// ---- POUs/POUs/FB/FB_Station05_Tear.TcPOU
FUNCTION_BLOCK FB_Station05_Tear EXTENDS FB_RollerConveyor
// =============================================================
// STACJA 5 - TEST WYTRZYMALOSCI NA ROZRYWANIE
// =============================================================
//
// Transporter rolkowy plus mechanika testu: blokada punktu
// zatrzymania, podnoszone szczeki chwytajace dolne deski
// i szesc silownikow rozrywajacych napierajacych na deski gorne.
//
// -------------------------------------------------------------
// DLACZEGO NIE MA PRZEJAZDU BEZ ZATRZYMANIA
// -------------------------------------------------------------
// Blokada stoi dokladnie w punkcie zatrzymania. Zeby przepuscic
// palete bez postoju, trzeba by ja opuscic ZANIM paleta dojedzie,
// czyli podjac decyzje na podstawie stanu, ktory dopiero ma
// nastapic. Blad w tej decyzji to paleta wjezdzajaca w podniesiona
// blokade z pelna predkoscia.
//
// Dlatego stacja 5 zatrzymuje KAZDA palete, takze odrzucona
// i takze przy wylaczonym tescie - wtedy sekwencja sprowadza sie
// do opuszczenia blokady. W GVL_PERSIST.aConv[5].Cfg nalezy
// ustawic xAllowPassThrough := FALSE.
//
// -------------------------------------------------------------
// KIEDY PODNOSI SIE BLOKADA
// -------------------------------------------------------------
// W chwili, gdy z poprzedniej stacji RUSZA paleta - czyli
// w M_BeginInfeed. Wtedy droga jest wolna na pewno, a czasu na
// ruch jest tyle, ile trwa przejazd miedzy stacjami.
//
// Podnoszenie jej czasowka po zjezdzie poprzedniej palety
// byloby zgadywaniem, czy paleta zeszla juz z blokady.
//
// -------------------------------------------------------------
// PRZEBIEG TESTU
// -------------------------------------------------------------
//   10  czasowka od potwierdzenia palety na blokadzie
//   20  podniesienie szczek
//   30  zamkniecie szczek (3 pary)
//   40  czasowka przed rozrywaniem
//   50  rozrywanie - kazdy silownik badany OSOBNO
//   60  otwarcie szczek
//   70  opuszczenie szczek
//   80  opuszczenie blokady
//   90  koniec
//
// Kazdy silownik rozrywajacy ma wlasny licznik czasu trzymania
// nacisku, bo wszystkie ida z inna predkoscia. Przekroczenie
// progu polozenia = deska odpadla: paleta staje sie NOK i nie
// przechodzi juz zadnych dalszych testow ani etykietowania.
VAR_INPUT

	stIn	: ST_St05_In;

END_VAR
VAR_OUTPUT

	stOut	: ST_St05_Out;

	// Krok sekwencji testu - do podgladu na HMI
	nTestStep		: INT;

	// Ktorego silownika rozrywajacego jeszcze czekamy (0 = zaden)
	nWaitPull		: INT;

	// Wynik dla biezacej palety
	axBoardBroken	: ARRAY[1..6] OF BOOL;

	// Wolna droga dla wjazdu: szczeki otwarte i opuszczone,
	// silowniki rozrywajace wycofane. Blokada NIE jest tu
	// warunkiem - podnosi sie dopiero w chwili wjazdu.
	xEntryReady		: BOOL;

	// Pelne polozenie spoczynkowe, z blokada w gorze
	xHomePosition	: BOOL;

	// Pierwszy silownik zglaszajacy blad i jego przyczyna.
	// nFaultyCyl: 1..3 szczeki, 4 blokada, 5 podnoszenie szczek,
	//             6..11 silowniki rozrywajace 1..6
	nFaultyCyl		: INT;
	eCylAlarm		: E_CylAlarm;

END_VAR
VAR

	pSt				: POINTER TO ST_St05Cfg;

	// Blokada punktu zatrzymania
	fbBlock			: FB_Cylinder;

	// Podnoszenie i opuszczanie szczek
	fbJawLift		: FB_Cylinder;

	// Szczeki - trzy pary, kazda para jeden zawor
	fbJaw			: ARRAY[1..3] OF FB_Cylinder;

	// Silowniki rozrywajace, indeksowane NUMEREM SILOWNIKA
	fbPull			: ARRAY[1..6] OF FB_Cylinder;

	axPullDone		: ARRAY[1..6] OF BOOL;

	tonSeq			: TON;
	tonOpWd			: TON;

	i				: INT;
	xAllJawsOpen	: BOOL;
	xAllJawsClosed	: BOOL;
	xAllPullBack	: BOOL;

END_VAR
VAR CONSTANT

	ST5_IDLE			: INT := 0;
	ST5_DELAY			: INT := 10;
	ST5_JAWLIFT_UP		: INT := 20;
	ST5_JAWS_CLOSE		: INT := 30;
	ST5_SETTLE			: INT := 40;
	ST5_PULL			: INT := 50;
	ST5_JAWS_OPEN		: INT := 60;
	ST5_JAWLIFT_DOWN	: INT := 70;
	ST5_BLOCK_DOWN		: INT := 80;
	ST5_DONE			: INT := 90;

END_VAR

// =============================================================
// CYKL STACJI 5
// =============================================================


// 1. Odswiezenie sprzezen silownikow.
//    Robimy to PRZED sekwencja, zeby decyzja "deska odpadla"
//    zapadala na swiezym odczycie przetwornika.
M_CallCylinders();


// 2. Warstwa transportu - wola M_OperationRequired
//    i M_OperationCycle
SUPER^();


// 3. Sprowadzenie mechaniki do polozenia spoczynkowego,
//    gdy stacja jest pusta
M_HomeCycle();


// 4. Przepisanie cewek na strukture wyjsciowa
M_MapOutputs();

METHOD PUBLIC M_ConfigStation
// Podpiecie nastaw stacji i wszystkich silownikow.
// Wolac raz, przy starcie, PO M_Config klasy bazowej.
VAR_INPUT
	pStCfg		: POINTER TO ST_St05Cfg;

	// Tablica rekordow silownikow - ADR(GVL_PERSIST.aCyl)
	pCylArray	: POINTER TO ARRAY[1..32] OF ST_CylPersist;

	// Pierwszy indeks przydzielony stacji. Stacja zajmuje
	// 11 kolejnych rekordow: szczeki 1..3, blokada,
	// podnoszenie szczek, silowniki rozrywajace 1..6.
	nCylBase	: INT;
END_VAR
VAR
	j			: INT;
END_VAR
pSt := pStCfg;

IF pCylArray = 0 THEN
	RETURN;
END_IF


// Szczeki
FOR j := 1 TO 3 DO
	fbJaw[j].M_Config(
		nId			:= nCylBase + j - 1,
		pPersist	:= ADR(pCylArray^[nCylBase + j - 1])
	);
END_FOR

// Blokada punktu zatrzymania
fbBlock.M_Config(
	nId			:= nCylBase + 3,
	pPersist	:= ADR(pCylArray^[nCylBase + 3])
);

// Podnoszenie szczek
fbJawLift.M_Config(
	nId			:= nCylBase + 4,
	pPersist	:= ADR(pCylArray^[nCylBase + 4])
);

// Silowniki rozrywajace
FOR j := 1 TO 6 DO
	fbPull[j].M_Config(
		nId			:= nCylBase + 4 + j,
		pPersist	:= ADR(pCylArray^[nCylBase + 4 + j])
	);
END_FOR
END_METHOD

METHOD PROTECTED M_CallCylinders
// Wywolanie wszystkich silownikow z ich sygnalami wejsciowymi
// oraz zebranie zbiorczych warunkow mechaniki.
VAR
	j	: INT;
END_VAR
fbBlock(
	eMode		:= eMode,
	xSafetyOK	:= xSafetyOK,
	xSwExtRaw	:= stIn.xBlockUpSw,
	xSwRetRaw	:= stIn.xBlockDownSw
);

fbJawLift(
	eMode		:= eMode,
	xSafetyOK	:= xSafetyOK,
	xSwExtRaw	:= stIn.xJawLiftUpSw,
	xSwRetRaw	:= stIn.xJawLiftDownSw
);


// Para szczek jest otwarta dopiero gdy OBA silowniki
// zglaszaja otwarcie
xAllJawsOpen	:= TRUE;
xAllJawsClosed	:= TRUE;

FOR j := 1 TO 3 DO

	fbJaw[j](
		eMode		:= eMode,
		xSafetyOK	:= xSafetyOK,
		xSwExtRaw	:= FALSE,
		xSwRetRaw	:= stIn.axJawOpenSw[j, 1] AND stIn.axJawOpenSw[j, 2]
	);

	IF NOT fbJaw[j].xRetracted THEN
		xAllJawsOpen := FALSE;
	END_IF

	IF NOT fbJaw[j].xExtended THEN
		xAllJawsClosed := FALSE;
	END_IF

END_FOR


xAllPullBack := TRUE;

FOR j := 1 TO 6 DO

	fbPull[j](
		eMode		:= eMode,
		xSafetyOK	:= xSafetyOK,
		diPosRaw	:= stIn.adiPullPos[j]
	);

	IF NOT fbPull[j].xRetracted THEN
		xAllPullBack := FALSE;
	END_IF

END_FOR


// Wolna droga dla wjazdu. Blokada nie jest tu warunkiem -
// podnosi sie dopiero wtedy, gdy z poprzedniej stacji rusza
// paleta, wiec przy pustej stacji stoi w dole.
xEntryReady := fbJawLift.xRetracted AND xAllJawsOpen AND xAllPullBack;

xHomePosition := xEntryReady AND fbBlock.xExtended;


M_ScanCylinderFaults();
END_METHOD

METHOD PROTECTED M_MapOutputs
VAR
	j	: INT;
END_VAR
stOut.xBlockExtend		:= fbBlock.xCoilExtend;
stOut.xBlockRetract		:= fbBlock.xCoilRetract;

stOut.xJawLiftExtend	:= fbJawLift.xCoilExtend;
stOut.xJawLiftRetract	:= fbJawLift.xCoilRetract;

FOR j := 1 TO 3 DO
	stOut.axJawClose[j] := fbJaw[j].xCoilExtend;
END_FOR

FOR j := 1 TO 6 DO
	stOut.axPullUp[j]	:= fbPull[j].xCoilExtend;
	stOut.axPullDown[j]	:= fbPull[j].xCoilRetract;
END_FOR
END_METHOD

METHOD PROTECTED M_HomeCycle
// Sprowadzenie mechaniki do polozenia gotowosci, gdy stacja
// jest pusta: szczeki otwarte i opuszczone, silowniki
// rozrywajace wycofane.
//
// BLOKADY TU NIE RUSZAMY. Podnosi sie dopiero w chwili, gdy
// z poprzedniej stacji rusza paleta - patrz M_BeginInfeed.
// Podnoszenie jej na czasowke po zjezdzie poprzedniej palety
// oznaczaloby zgadywanie, czy paleta zeszla juz z blokady.
//
// Poza stanem pustym komendy zostaja takie, jakie zostawila
// sekwencja testu.
VAR
	j	: INT;
END_VAR
IF (eState <> NODE_EMPTY) AND (eState <> NODE_INIT) THEN
	RETURN;
END_IF

fbJawLift.M_Retract();

FOR j := 1 TO 3 DO
	fbJaw[j].M_Retract();
END_FOR

FOR j := 1 TO 6 DO
	fbPull[j].M_Retract();
END_FOR
END_METHOD

METHOD PUBLIC M_BeginInfeed
// Poprzednia stacja wlasnie ruszyla z paleta.
//
// To jest moment na podniesienie blokady: droga jest wolna,
// paleta dopiero wjezdza, a czasu na ruch jest tyle, ile trwa
// przejazd miedzy stacjami. Nie zgadujemy niczego czasowka.
VAR_INPUT
	pSource		: POINTER TO FB_TransportNodeBase;
	xNok		: BOOL;
	nLoadId		: UDINT;
END_VAR
SUPER^.M_BeginInfeed(
	pSource	:= pSource,
	xNok	:= xNok,
	nLoadId	:= nLoadId
);

fbBlock.M_Extend();
END_METHOD

METHOD PROTECTED M_ScanCylinderFaults
// Pierwszy silownik w bledzie zostaje wskazany na wyjsciu,
// a stacja idzie w alarm. Kolejne go nie nadpisuja - operator
// ma zobaczyc przyczyne, nie skutek.
VAR
	j	: INT;
END_VAR
IF nFaultyCyl <> 0 THEN
	RETURN;
END_IF

FOR j := 1 TO 3 DO
	IF fbJaw[j].xAlarm AND (nFaultyCyl = 0) THEN
		nFaultyCyl	:= j;
		eCylAlarm	:= fbJaw[j].eAlarm;
	END_IF
END_FOR

IF fbBlock.xAlarm AND (nFaultyCyl = 0) THEN
	nFaultyCyl	:= 4;
	eCylAlarm	:= fbBlock.eAlarm;
END_IF

IF fbJawLift.xAlarm AND (nFaultyCyl = 0) THEN
	nFaultyCyl	:= 5;
	eCylAlarm	:= fbJawLift.eAlarm;
END_IF

FOR j := 1 TO 6 DO
	IF fbPull[j].xAlarm AND (nFaultyCyl = 0) THEN
		nFaultyCyl	:= 5 + j;
		eCylAlarm	:= fbPull[j].eAlarm;
	END_IF
END_FOR

IF nFaultyCyl <> 0 THEN
	M_RaiseAlarm(eNew := ALM_OPERATION_FAILED);
END_IF
END_METHOD

METHOD PUBLIC M_WhyCannotAccept : E_WaitCause
// Warunki klasy bazowej plus wlasne: paleta nie ma prawa
// wjechac, dopoki blokada nie stoi w gorze, a szczeki nie sa
// otwarte i opuszczone.
M_WhyCannotAccept := SUPER^.M_WhyCannotAccept();

IF M_WhyCannotAccept <> WAIT_NONE THEN
	RETURN;
END_IF

IF NOT xEntryReady THEN
	M_WhyCannotAccept := WAIT_STATION_NOT_READY;
END_IF
END_METHOD

METHOD PROTECTED M_OperationRequired : BOOL
// Zawsze TRUE. Nawet paleta odrzucona i nawet przy wylaczonym
// tescie musi sie tu zatrzymac - blokada stoi w punkcie
// zatrzymania i trzeba ja opuscic, zanim paleta pojedzie dalej.
M_OperationRequired := TRUE;
END_METHOD

METHOD PROTECTED M_TestEnabled : BOOL
// Czy dla tej palety w ogole robimy test.
M_TestEnabled := FALSE;

IF pP = 0 THEN
	RETURN;
END_IF

// Operator wylaczyl stacje
IF NOT pP^.Cfg.xStationEnabled THEN
	RETURN;
END_IF

// Paleta juz odrzucona - zadnych dalszych testow
IF pP^.Mem.xLoadNok THEN
	RETURN;
END_IF

M_TestEnabled := TRUE;
END_METHOD

METHOD PROTECTED M_OperationCycle : BOOL
// Sekwencja stacji. Zwraca TRUE, gdy paleta moze jechac dalej.
VAR
	j	: INT;
END_VAR
M_OperationCycle := FALSE;

IF pSt = 0 THEN
	M_RaiseAlarm(eNew := ALM_NOT_CONFIGURED);
	RETURN;
END_IF


// ---------------------------------------------------------
// WATCHDOG CALEJ OPERACJI
// ---------------------------------------------------------

tonOpWd(IN := (nTestStep <> ST5_IDLE), PT := pSt^.tOpWatchdog);

IF tonOpWd.Q THEN
	M_RaiseAlarm(eNew := ALM_OPERATION_FAILED);
	RETURN;
END_IF


CASE nTestStep OF

ST5_IDLE:
	// Start operacji dla nowej palety
	nWaitPull := 0;

	FOR j := 1 TO 6 DO
		axBoardBroken[j]	:= FALSE;
		axPullDone[j]		:= FALSE;
	END_FOR

	tonSeq(IN := FALSE);

	IF M_TestEnabled() THEN
		nTestStep := ST5_DELAY;
	ELSE
		// Bez testu idziemy przez wycofywanie mechaniki, a nie
		// prosto do blokady. Przy pustej stacji te kroki mijaja
		// natychmiast, ale gdy test zostal przerwany w polowie
		// i paleta stala sie NOK - szczeki i silowniki moga byc
		// w dowolnym polozeniu i trzeba je najpierw sciagnac.
		nTestStep := ST5_JAWS_OPEN;
	END_IF


ST5_DELAY:
	tonSeq(IN := TRUE, PT := pSt^.tDetectToLift);

	IF tonSeq.Q THEN
		tonSeq(IN := FALSE);
		nTestStep := ST5_JAWLIFT_UP;
	END_IF


ST5_JAWLIFT_UP:
	fbJawLift.M_Extend();

	IF fbJawLift.xExtended THEN
		nTestStep := ST5_JAWS_CLOSE;
	END_IF


ST5_JAWS_CLOSE:
	FOR j := 1 TO 3 DO
		fbJaw[j].M_Extend();
	END_FOR

	IF xAllJawsClosed THEN
		nTestStep := ST5_SETTLE;
	END_IF


ST5_SETTLE:
	tonSeq(IN := TRUE, PT := pSt^.tJawsToPull);

	IF tonSeq.Q THEN
		tonSeq(IN := FALSE);
		nTestStep := ST5_PULL;
	END_IF


ST5_PULL:
	M_PullCycle();

	IF xAllPullBack AND (nWaitPull = 0) THEN
		nTestStep := ST5_JAWS_OPEN;
	END_IF


ST5_JAWS_OPEN:
	// Silowniki rozrywajace sciagamy takze tutaj - tedy prowadzi
	// droga wyjscia z przerwanego testu
	FOR j := 1 TO 6 DO
		fbPull[j].M_Retract();
	END_FOR

	FOR j := 1 TO 3 DO
		fbJaw[j].M_Retract();
	END_FOR

	IF xAllJawsOpen AND xAllPullBack THEN
		nTestStep := ST5_JAWLIFT_DOWN;
	END_IF


ST5_JAWLIFT_DOWN:
	fbJawLift.M_Retract();

	IF fbJawLift.xRetracted THEN
		nTestStep := ST5_BLOCK_DOWN;
	END_IF


ST5_BLOCK_DOWN:
	fbBlock.M_Retract();

	IF fbBlock.xRetracted THEN
		nTestStep := ST5_DONE;
	END_IF


ST5_DONE:
	// Wyjazd dozwolony dopiero gdy WSZYSTKO jest wycofane
	IF NOT xAllJawsOpen THEN
		RETURN;
	END_IF

	IF NOT fbJawLift.xRetracted THEN
		RETURN;
	END_IF

	IF NOT xAllPullBack THEN
		RETURN;
	END_IF

	IF NOT fbBlock.xRetracted THEN
		RETURN;
	END_IF

	tonOpWd(IN := FALSE);
	nTestStep			:= ST5_IDLE;
	M_OperationCycle	:= TRUE;


ELSE
	nTestStep := ST5_IDLE;

END_CASE
END_METHOD

METHOD PROTECTED M_PullCycle
// Rozrywanie. Kazdy silownik prowadzony OSOBNO - maja rozne
// predkosci, wiec kazdy dochodzi do progu w innej chwili
// i kazdy ma wlasny licznik czasu trzymania nacisku.
VAR
	j	: INT;
END_VAR
nWaitPull := 0;

FOR j := 1 TO 6 DO

	M_PullOne(j := j);

	IF NOT axPullDone[j] THEN
		nWaitPull := j;
	END_IF

END_FOR
END_METHOD

METHOD PROTECTED M_PullOne
// Jeden silownik rozrywajacy.
//
// Kolejnosc warunkow jest istotna: najpierw sprawdzamy, czy
// deska odpadla, i dopiero potem czy nacisk zostal utrzymany.
// Odwrotnie mozna by uznac za dobra deske, ktora wlasnie pekla.
VAR_INPUT
	j	: INT;
END_VAR
// Ten juz zbadany - wraca do bazy
IF axPullDone[j] THEN
	fbPull[j].M_Retract();
	RETURN;
END_IF


// Wysunal sie dalej, niz moglby z cala paleta - deska odpadla
IF fbPull[j].xOverLimit THEN
	axBoardBroken[j]	:= TRUE;
	axPullDone[j]		:= TRUE;

	IF pP <> 0 THEN
		pP^.Mem.xLoadNok	:= TRUE;
		xPersistDirty		:= TRUE;
	END_IF

	fbPull[j].M_Retract();
	RETURN;
END_IF


// Nacisk utrzymany przez nastawiony czas - deska wytrzymala
IF fbPull[j].xHoldDone THEN
	axPullDone[j] := TRUE;
	fbPull[j].M_Retract();
	RETURN;
END_IF


fbPull[j].M_Extend();
END_METHOD

METHOD PUBLIC M_Reset : BOOL
VAR
	j	: INT;
END_VAR
fbBlock.M_Reset();
fbJawLift.M_Reset();

FOR j := 1 TO 3 DO
	fbJaw[j].M_Reset();
END_FOR

FOR j := 1 TO 6 DO
	fbPull[j].M_Reset();
END_FOR

tonSeq(IN := FALSE);
tonOpWd(IN := FALSE);

nTestStep	:= ST5_IDLE;
nWaitPull	:= 0;
nFaultyCyl	:= 0;
eCylAlarm	:= ALM_CYL_NONE;

M_Reset := SUPER^.M_Reset();
END_METHOD

METHOD PUBLIC M_ManCylinder
// Sterowanie reczne pojedynczym silownikiem stacji.
// nSel: 1..3 szczeki, 4 blokada, 5 podnoszenie szczek,
//       6..11 silowniki rozrywajace 1..6
VAR_INPUT
	nSel	: INT;
	xExt	: BOOL;
	xRet	: BOOL;
END_VAR
IF (nSel >= 1) AND (nSel <= 3) THEN
	fbJaw[nSel].M_ManJog(xExt := xExt, xRet := xRet);
	RETURN;
END_IF

IF nSel = 4 THEN
	fbBlock.M_ManJog(xExt := xExt, xRet := xRet);
	RETURN;
END_IF

IF nSel = 5 THEN
	fbJawLift.M_ManJog(xExt := xExt, xRet := xRet);
	RETURN;
END_IF

IF (nSel >= 6) AND (nSel <= 11) THEN
	fbPull[nSel - 5].M_ManJog(xExt := xExt, xRet := xRet);
END_IF
END_METHOD

METHOD PUBLIC M_ZeroPull : BOOL
// Bazowanie przetwornikow silownikow rozrywajacych.
// Zero jest na silowniku WYCOFANYM, bez palety.
// nSel = 0 zeruje wszystkie naraz.
VAR_INPUT
	nSel	: INT;
END_VAR
VAR
	j		: INT;
END_VAR
M_ZeroPull := FALSE;

IF nSel = 0 THEN
	FOR j := 1 TO 6 DO
		fbPull[j].M_Zero();
	END_FOR
	M_ZeroPull := TRUE;
	RETURN;
END_IF

IF (nSel < 1) OR (nSel > 6) THEN
	RETURN;
END_IF

M_ZeroPull := fbPull[nSel].M_Zero();
END_METHOD

END_FUNCTION_BLOCK

// ---- POUs/POUs/FB/FB_StationPickup.TcPOU
FUNCTION_BLOCK FB_StationPickup EXTENDS FB_RollerConveyor
// =============================================================
// STACJA ODBIORU - 13 (stosy dobre) I 16 (palety odrzucone)
// =============================================================
//
// Koniec drogi: ladunek stoi na czujnikach i zabiera go operator.
// Nie ma nastepnika, wiec zwolnienie miejsca musi wykryc sama
// stacja.
//
// Dwa sposoby, przelaczane nastawa Cfg.xPickupByButton:
//
//   TRUE  - operator potwierdza przyciskiem. Sprawdzamy wtedy,
//           czy ladunek faktycznie zniknal z czujnikow. Jesli
//           nie zniknal, nie robimy nic - przycisk nie jest
//           dowodem na to, ze cos zostalo zabrane.
//
//   FALSE - miejsce uznajemy za wolne po Cfg.tPickupTimeout
//           od zniknieca ladunku z czujnikow.
VAR_INPUT

	// Przycisk operatora "zabralem"
	xPickupButton	: BOOL;

END_VAR
VAR_OUTPUT

	// Czeka na odbior
	xWaitingPickup	: BOOL;

END_VAR
VAR

	tonPickup	: TON;
	rtrgButton	: R_TRIG;

END_VAR

SUPER^();

M_PickupCycle();

METHOD PROTECTED M_PickupCycle
VAR
	xFree	: BOOL;
END_VAR
xWaitingPickup := FALSE;

IF pP = 0 THEN
	RETURN;
END_IF

IF NOT pP^.Mem.xLoadPresent THEN
	tonPickup(IN := FALSE);
	rtrgButton(CLK := xPickupButton);
	RETURN;
END_IF

xWaitingPickup	:= TRUE;
eWait			:= WAIT_PICKUP;


// Pole czujnikow wolne. Przy wylaczonych czujnikach nie mamy
// czym tego stwierdzic - wtedy decyduje sam przycisk.
IF xSensUsable THEN
	xFree := xSensLoadNone;
ELSE
	xFree := TRUE;
END_IF


// --- potwierdzenie przyciskiem ---
IF pP^.Cfg.xPickupByButton THEN

	rtrgButton(CLK := xPickupButton);

	IF NOT rtrgButton.Q THEN
		RETURN;
	END_IF

	// Przycisk wcisniety, ale ladunek dalej lezy - nic nie robimy
	IF NOT xFree THEN
		RETURN;
	END_IF

	M_ClearLoad();
	RETURN;

END_IF


// --- odliczanie od zniknieca z czujnikow ---
rtrgButton(CLK := xPickupButton);

tonPickup(IN := xFree, PT := pP^.Cfg.tPickupTimeout);

IF tonPickup.Q THEN
	tonPickup(IN := FALSE);
	M_ClearLoad();
END_IF
END_METHOD

METHOD PROTECTED M_OperationRequired : BOOL
// Nie ma operacji technologicznej - ladunek po prostu czeka.
M_OperationRequired := FALSE;
END_METHOD

END_FUNCTION_BLOCK

// ---- POUs/PRG_Machine.TcPOU
PROGRAM PRG_Machine
// =============================================================
// TESTER PALET - PELNA APLIKACJA (CHWILOWO NIEWYWOLYWANA)
// =============================================================
//
// Ten program NIE jest wolany z zadania. MAIN wykonuje teraz
// wylacznie test ruchu transporterow. Zeby wrocic do pelnej
// aplikacji, wystarczy w MAIN wywolac PRG_Machine() zamiast
// akcji testowych.
// =============================================================
// =============================================================
//
// Wszystkie bity, ktore trzeba podlinkowac albo przestawiac
// online, siedza W TYM PROGRAMIE, na gorze deklaracji. Nie
// trzeba ich szukac po blokach.
//
// -------------------------------------------------------------
// CZYM SIE ROZNI OD WERSJI DOCELOWEJ
// -------------------------------------------------------------
//   - czujniki pracuja w logice WPROST: 1 = jest paleta
//     (docelowo bedzie odwrotnie, przelacza to jeden bit
//     w nastawach kazdej stacji)
//   - stacje bez czujnikow jada na czasowki
//   - silowniki nie maja czujnikow polozenia - kazdy ruch
//     jest potwierdzany czasowka
//   - czestotliwosc wszystkich falownikow 15 Hz
//   - przejazd bez zatrzymania wylaczony na wszystkich stacjach
//   - werdykt OK / NOK wystawia licznik: co piata paleta NOK
//
// ACT_Config nadpisuje nastawy nieulotne przy kazdym starcie
// sterownika. W wersji docelowej ta akcja znika i nastawy
// zostaja pod kontrola operatora.
VAR

	// =========================================================
	// 1. STEROWANIE - DO ZMIANY ONLINE
	// =========================================================

	// Tryb pracy maszyny
	eMode				: E_MachineMode := MODE_AUTO;

	// Zezwolenie z lancucha bezpieczenstwa.
	// Na czas uruchomienia mozna trzymac TRUE z palca.
	xSafetyOK			: BOOL := TRUE;

	// RECZNE ZEZWOLENIE NA PRZEJAZDY MIEDZY STACJAMI.
	// FALSE zatrzymuje wydawanie ladunkow - maszyna stoi tam,
	// gdzie jest, i nic sie nie przesuwa dalej.
	xTransferEnable		: BOOL := TRUE;

	// Operator wstawil stos na stacje 1.
	// Czujnik stacji 1 nie widzi stosu, wiec informacje
	// podajemy tym bitem - dziala na zbocze.
	xCmdStackInserted	: BOOL;

	// Kasowanie alarmow wszystkich stacji - zbocze
	xCmdReset			: BOOL;

	// RESET MASZYNY DO STANU ZEROWEGO - zbocze.
	// Kasuje pamiec obecnosci na wszystkich stacjach oraz
	// liczniki desztaplarki i sztaplarki. Do uzycia, gdy
	// maszyne trzeba oproznic recznie.
	xCmdClearMachine	: BOOL;


	// =========================================================
	// 2. CZUJNIKI - DO PODLINKOWANIA
	// =========================================================
	//
	// Logika WPROST: 0 = nie ma palety, 1 = jest paleta.

	xSens_St01			: BOOL;		// stacja 1
	xSens_St03			: BOOL;		// stacja 3
	xSens_St04_Entry	: BOOL;		// stacja 4 - wjazd palety
	xSens_St04_Stop		: BOOL;		// stacja 4 - pozycja koncowa
	xSens_St07			: BOOL;		// stacja 7
	xSens_St11			: BOOL;		// stacja 11
	xSens_St13			: BOOL;		// stacja 13
	xSens_St16			: BOOL;		// stacja 16

	// Enkodery absolutne wozkow. Pozycje robocze wpisujemy
	// z palca w ACT_Config - patrz sekcja DESZTAPLARKA.
	diEnc_St03			: DINT;
	diEnc_St11			: DINT;


	// =========================================================
	// 3. WYJSCIA SZCZEK - DO PODLINKOWANIA
	// =========================================================

	xOut_St03_JawClose	: BOOL;
	xOut_St03_JawOpen	: BOOL;
	xOut_St11_JawClose	: BOOL;
	xOut_St11_JawOpen	: BOOL;


	// =========================================================
	// 4. STACJE
	// =========================================================

	fbSt01	: FB_RollerConveyor;
	fbSt02	: FB_RollerConveyor;
	fbSt03	: FB_Station03_Destack;
	fbSt04	: FB_Station04_Press;
	fbSt05	: FB_Station05_Tear;
	fbSt06	: FB_RollerConveyor;
	fbSt07	: FB_RollerConveyor;
	fbSt08	: FB_RollerConveyor;
	fbSt09	: FB_RollerConveyor;
	fbSt10	: FB_RollerConveyor;
	fbSt11	: FB_Station11_Stack;
	fbSt12	: FB_RollerConveyor;
	fbSt13	: FB_StationPickup;
	fbSt14	: FB_RollerConveyor;
	fbSt15	: FB_RollerConveyor;
	fbSt16	: FB_StationPickup;

	// Wskazniki na wezly - do podpinania sasiadow i do resetu
	aNode	: ARRAY[1..16] OF POINTER TO FB_TransportNodeBase;


	// =========================================================
	// 5. NAPEDY
	// =========================================================

	fbNord	: ARRAY[1..20] OF FB_NordSK550PP;

	// Lustro diagnostyczne napedow
	aeDrvState		: ARRAY[1..20] OF E_NordSK550P_State;
	axDrvRunning	: ARRAY[1..20] OF BOOL;
	axDrvError		: ARRAY[1..20] OF BOOL;
	alrDrvFreqAct	: ARRAY[1..20] OF LREAL;


	// =========================================================
	// 6. DIAGNOSTYKA STACJI - PODGLAD ONLINE
	// =========================================================

	aeState		: ARRAY[1..16] OF E_NodeState;
	aeWait		: ARRAY[1..16] OF E_WaitCause;
	aeAlarm		: ARRAY[1..16] OF E_NodeAlarm;
	axOccupied	: ARRAY[1..16] OF BOOL;
	axNok		: ARRAY[1..16] OF BOOL;

	// Licznik palet i werdykty
	nPalletsDone	: INT;
	nOkCount		: INT;
	nNokCount		: INT;


	// =========================================================
	// 7. WEWNETRZNE
	// =========================================================

	xInit		: BOOL;
	i			: INT;

	rtrgStack	: R_TRIG;
	rtrgReset	: R_TRIG;
	rtrgClear	: R_TRIG;
	rtrgSt05	: R_TRIG;

	nLoadSeq	: UDINT;

END_VAR
VAR CONSTANT

	// P105 falownikow
	cFmax		: LREAL := 50.0;

	// Liczba falownikow zmapowanych w .tsproj
	cNumDrives	: INT := 19;

	// Czestotliwosc robocza wersji testowej
	cTestFreq	: LREAL := 15.0;

	// Co ktora paleta ma byc uznana za NOK
	cNokEvery	: INT := 5;

END_VAR

// =============================================================
// MAIN - TESTER PALET
// =============================================================
//
// Kolejnosc jest czescia kontraktu: najpierw stacje, bo wolaja
// metody blokow napedu, dopiero potem same napedy.


// Jednorazowa konfiguracja
ACT_Config();

// Komendy operatora
ACT_Commands();

// Stacje
ACT_Stations();

// Test: werdykt OK / NOK i trasowanie na stacji 8
ACT_Verdict();

// Napedy
ACT_Drives();

// Podglad
ACT_Diag();

ACTION ACT_Config:
// =============================================================
// ACT_Config
// Konfiguracja jednorazowa - WERSJA TESTOWA
// =============================================================
//
// Ta akcja NADPISUJE nastawy nieulotne przy kazdym starcie
// sterownika. Tak ma byc na czas uruchomienia: chcemy miec
// pewnosc, od czego zaczynamy. W wersji docelowej ta akcja
// znika, a nastawy zostaja pod kontrola operatora.

IF xInit THEN
	RETURN;
END_IF

xInit := TRUE;


// -------------------------------------------------------------
// WSKAZNIKI NA WEZLY
// -------------------------------------------------------------

aNode[1]  := ADR(fbSt01);
aNode[2]  := ADR(fbSt02);
aNode[3]  := ADR(fbSt03);
aNode[4]  := ADR(fbSt04);
aNode[5]  := ADR(fbSt05);
aNode[6]  := ADR(fbSt06);
aNode[7]  := ADR(fbSt07);
aNode[8]  := ADR(fbSt08);
aNode[9]  := ADR(fbSt09);
aNode[10] := ADR(fbSt10);
aNode[11] := ADR(fbSt11);
aNode[12] := ADR(fbSt12);
aNode[13] := ADR(fbSt13);
aNode[14] := ADR(fbSt14);
aNode[15] := ADR(fbSt15);
aNode[16] := ADR(fbSt16);


// -------------------------------------------------------------
// NASTAWY WSPOLNE
// -------------------------------------------------------------

FOR i := 1 TO 16 DO

	GVL_PERSIST.aConv[i].Cfg.lrFreqAuto			:= cTestFreq;
	GVL_PERSIST.aConv[i].Cfg.lrFreqManual		:= cTestFreq;
	GVL_PERSIST.aConv[i].Cfg.tStopDelay			:= T#150MS;

	// Wersja testowa: 1 = jest paleta
	GVL_PERSIST.aConv[i].Cfg.xSensorsInverted	:= FALSE;

	GVL_PERSIST.aConv[i].Cfg.tSensorSettle		:= T#1S;
	GVL_PERSIST.aConv[i].Cfg.tInfeedWatchdog	:= T#40S;
	GVL_PERSIST.aConv[i].Cfg.tOutfeedWatchdog	:= T#40S;
	GVL_PERSIST.aConv[i].Cfg.tBlindTravel		:= T#5S;
	GVL_PERSIST.aConv[i].Cfg.tClearDelay		:= T#500MS;

	GVL_PERSIST.aConv[i].Cfg.xStationEnabled	:= TRUE;
	GVL_PERSIST.aConv[i].Cfg.nResumeRetries		:= 1;

	// Na czas uruchomienia kazda paleta zatrzymuje sie na
	// kazdej stacji - latwiej obserwowac
	GVL_PERSIST.aConv[i].Cfg.xAllowPassThrough	:= FALSE;

	// Domyslnie oba czujniki wylaczone, czyli przejazd na
	// czasowke. Ponizej wlaczamy tylko te, ktore istnieja.
	GVL_PERSIST.aConv[i].Cfg.xSensor1Enabled	:= FALSE;
	GVL_PERSIST.aConv[i].Cfg.xSensor2Enabled	:= FALSE;
	GVL_PERSIST.aConv[i].Cfg.xInvertDirection	:= FALSE;

END_FOR


// -------------------------------------------------------------
// CZUJNIKI, KTORE ISTNIEJA
// -------------------------------------------------------------

GVL_PERSIST.aConv[3].Cfg.xSensor1Enabled	:= TRUE;
GVL_PERSIST.aConv[4].Cfg.xSensor1Enabled	:= TRUE;
GVL_PERSIST.aConv[7].Cfg.xSensor1Enabled	:= TRUE;
GVL_PERSIST.aConv[11].Cfg.xSensor1Enabled	:= TRUE;
GVL_PERSIST.aConv[13].Cfg.xSensor1Enabled	:= TRUE;
GVL_PERSIST.aConv[16].Cfg.xSensor1Enabled	:= TRUE;


// -------------------------------------------------------------
// ODWROCONY KIERUNEK - ZLE PODLACZONE SILNIKI
// -------------------------------------------------------------
//
// Stacje 1, 5, 6, 7, 8, 9, 14, 15, 16. Do poprawy w szafie,
// na razie odwracamy bit.

GVL_PERSIST.aConv[1].Cfg.xInvertDirection	:= TRUE;
GVL_PERSIST.aConv[5].Cfg.xInvertDirection	:= TRUE;
GVL_PERSIST.aConv[6].Cfg.xInvertDirection	:= TRUE;
GVL_PERSIST.aConv[7].Cfg.xInvertDirection	:= TRUE;
GVL_PERSIST.aConv[8].Cfg.xInvertDirection	:= TRUE;
GVL_PERSIST.aConv[9].Cfg.xInvertDirection	:= TRUE;
GVL_PERSIST.aConv[14].Cfg.xInvertDirection	:= TRUE;
GVL_PERSIST.aConv[15].Cfg.xInvertDirection	:= TRUE;
GVL_PERSIST.aConv[16].Cfg.xInvertDirection	:= TRUE;


// -------------------------------------------------------------
// CZASY PRZEJAZDU NA STACJACH BEZ CZUJNIKOW
// -------------------------------------------------------------

GVL_PERSIST.aConv[1].Cfg.tBlindTravel		:= T#4S;
GVL_PERSIST.aConv[2].Cfg.tBlindTravel		:= T#5S;
GVL_PERSIST.aConv[5].Cfg.tBlindTravel		:= T#5S;
GVL_PERSIST.aConv[6].Cfg.tBlindTravel		:= T#5S;
GVL_PERSIST.aConv[8].Cfg.tBlindTravel		:= T#5S;

// Transporter lancuchowy - przejazd poprzeczny
GVL_PERSIST.aConv[9].Cfg.tBlindTravel		:= T#6S;

GVL_PERSIST.aConv[10].Cfg.tBlindTravel		:= T#5S;
GVL_PERSIST.aConv[12].Cfg.tBlindTravel		:= T#5S;
GVL_PERSIST.aConv[14].Cfg.tBlindTravel		:= T#5S;
GVL_PERSIST.aConv[15].Cfg.tBlindTravel		:= T#5S;


// -------------------------------------------------------------
// ODBIOR PRZEZ OPERATORA - STACJE 13 I 16
// -------------------------------------------------------------
//
// Bez przycisku: miejsce jest wolne po 5 s od zniknieca
// ladunku z czujnika.

GVL_PERSIST.aConv[13].Cfg.xPickupByButton	:= FALSE;
GVL_PERSIST.aConv[13].Cfg.tPickupTimeout	:= T#5S;
GVL_PERSIST.aConv[16].Cfg.xPickupByButton	:= FALSE;
GVL_PERSIST.aConv[16].Cfg.tPickupTimeout	:= T#5S;


// -------------------------------------------------------------
// SILOWNIKI - BEZ CZUJNIKOW, RUCH NA CZASOWKI
// -------------------------------------------------------------

FOR i := 1 TO 32 DO
	GVL_PERSIST.aCyl[i].Cfg.eFeedback			:= CYLFB_NONE;
	GVL_PERSIST.aCyl[i].Cfg.eValve				:= CYLV_DOUBLE;
	GVL_PERSIST.aCyl[i].Cfg.xExtendFbEnabled	:= FALSE;
	GVL_PERSIST.aCyl[i].Cfg.xRetractFbEnabled	:= FALSE;
	GVL_PERSIST.aCyl[i].Cfg.xExtendWdEnabled	:= FALSE;
	GVL_PERSIST.aCyl[i].Cfg.xRetractWdEnabled	:= FALSE;
	GVL_PERSIST.aCyl[i].Cfg.tExtendDelay		:= T#0MS;
	GVL_PERSIST.aCyl[i].Cfg.tRetractDelay		:= T#0MS;
	GVL_PERSIST.aCyl[i].Cfg.tExtendSubst		:= T#3S;
	GVL_PERSIST.aCyl[i].Cfg.tRetractSubst		:= T#3S;
END_FOR

// Dociski stacji 4 - szybciej niz reszta
FOR i := 1 TO 3 DO
	GVL_PERSIST.aCyl[i].Cfg.tExtendSubst		:= T#1S;
	GVL_PERSIST.aCyl[i].Cfg.tRetractSubst		:= T#1S;
END_FOR

// Blokada stacji 5 - zawor 3-polozeniowy
GVL_PERSIST.aCyl[15].Cfg.eValve					:= CYLV_3POS_MID;

// Szczeki desztaplarki i sztaplarki - 5 s na ruch
GVL_PERSIST.aCyl[25].Cfg.tExtendSubst			:= T#5S;
GVL_PERSIST.aCyl[25].Cfg.tRetractSubst			:= T#5S;
GVL_PERSIST.aCyl[26].Cfg.tExtendSubst			:= T#5S;
GVL_PERSIST.aCyl[26].Cfg.tRetractSubst			:= T#5S;


// -------------------------------------------------------------
// STACJA 4
// -------------------------------------------------------------

GVL_PERSIST.St04.xPreSensorInstalled	:= TRUE;
GVL_PERSIST.St04.xPreSensorInverted		:= FALSE;
GVL_PERSIST.St04.tPreToUpper			:= T#1S200MS;
GVL_PERSIST.St04.tEntryToUpper			:= T#3S;
GVL_PERSIST.St04.tUpperToLower			:= T#400MS;
GVL_PERSIST.St04.tOpWatchdog			:= T#60S;
GVL_PERSIST.St04.lrRollerFreq			:= cTestFreq;


// -------------------------------------------------------------
// STACJA 5
// -------------------------------------------------------------

GVL_PERSIST.St05.tDetectToLift		:= T#500MS;
GVL_PERSIST.St05.tJawsToPull		:= T#500MS;
GVL_PERSIST.St05.tOpWatchdog		:= T#120S;


// -------------------------------------------------------------
// DESZTAPLARKA - POZYCJE Z PALCA
// -------------------------------------------------------------
//
// Wartosci do poprawienia po zmierzeniu na maszynie.
// Musza tworzyc ciag - kod to sprawdza.

GVL_PERSIST.St03.Cfg.diPosBottom		:= 1000;
GVL_PERSIST.St03.Cfg.diPosMiddle		:= 2000;
GVL_PERSIST.St03.Cfg.diPosTop			:= 3000;
GVL_PERSIST.St03.Cfg.diWindow			:= 20;
GVL_PERSIST.St03.Cfg.diSlowZone			:= 300;
GVL_PERSIST.St03.Cfg.xIncreaseIsForward	:= TRUE;
GVL_PERSIST.St03.Cfg.lrFreqFast			:= cTestFreq;
GVL_PERSIST.St03.Cfg.lrFreqSlow			:= cTestFreq;
GVL_PERSIST.St03.Cfg.lrFreqManual		:= cTestFreq;
GVL_PERSIST.St03.Cfg.tMoveWatchdog		:= T#30S;
GVL_PERSIST.St03.Cfg.tSettle			:= T#200MS;
GVL_PERSIST.St03.Cfg.nStackSize			:= 15;


// -------------------------------------------------------------
// SZTAPLARKA - POZYCJE Z PALCA, INNE NIZ DESZTAPLARKI
// -------------------------------------------------------------

GVL_PERSIST.St11.Cfg.diPosBottom		:= 5000;
GVL_PERSIST.St11.Cfg.diPosMiddle		:= 6000;
GVL_PERSIST.St11.Cfg.diPosTop			:= 7000;
GVL_PERSIST.St11.Cfg.diWindow			:= 20;
GVL_PERSIST.St11.Cfg.diSlowZone			:= 300;
GVL_PERSIST.St11.Cfg.xIncreaseIsForward	:= TRUE;
GVL_PERSIST.St11.Cfg.lrFreqFast			:= cTestFreq;
GVL_PERSIST.St11.Cfg.lrFreqSlow			:= cTestFreq;
GVL_PERSIST.St11.Cfg.lrFreqManual		:= cTestFreq;
GVL_PERSIST.St11.Cfg.tMoveWatchdog		:= T#30S;
GVL_PERSIST.St11.Cfg.tSettle			:= T#200MS;
GVL_PERSIST.St11.Cfg.nStackSize			:= 15;


// -------------------------------------------------------------
// PODPIECIE REKORDOW I NAPEDOW
// -------------------------------------------------------------

FOR i := 1 TO 16 DO
	aNode[i]^.M_Config(nId := i, pPersist := ADR(GVL_PERSIST.aConv[i]));
END_FOR

// Przydzial falownikow wg listy z dokumentacji
fbSt01.M_ConfigDrive(pDrv := ADR(fbNord[8]));
fbSt02.M_ConfigDrive(pDrv := ADR(fbNord[9]));
fbSt03.M_ConfigDrive(pDrv := ADR(fbNord[10]));
fbSt04.M_ConfigDrive(pDrv := ADR(fbNord[4]));
fbSt05.M_ConfigDrive(pDrv := ADR(fbNord[5]));
fbSt06.M_ConfigDrive(pDrv := ADR(fbNord[6]));
fbSt07.M_ConfigDrive(pDrv := ADR(fbNord[11]));
fbSt08.M_ConfigDrive(pDrv := ADR(fbNord[12]));
fbSt09.M_ConfigDrive(pDrv := ADR(fbNord[7]));
fbSt10.M_ConfigDrive(pDrv := ADR(fbNord[16]));
fbSt11.M_ConfigDrive(pDrv := ADR(fbNord[13]));
fbSt12.M_ConfigDrive(pDrv := ADR(fbNord[14]));
fbSt13.M_ConfigDrive(pDrv := ADR(fbNord[15]));
fbSt14.M_ConfigDrive(pDrv := ADR(fbNord[17]));
fbSt15.M_ConfigDrive(pDrv := ADR(fbNord[18]));
fbSt16.M_ConfigDrive(pDrv := ADR(fbNord[19]));


// Stacja 4 - rolki dociskowe na falowniku 3
fbSt04.M_ConfigStation(
	pStCfg		:= ADR(GVL_PERSIST.St04),
	pRollerDrv	:= ADR(fbNord[3]),
	pCylArray	:= ADR(GVL_PERSIST.aCyl),
	nCylBase	:= 1
);

// Stacja 5
fbSt05.M_ConfigStation(
	pStCfg		:= ADR(GVL_PERSIST.St05),
	pCylArray	:= ADR(GVL_PERSIST.aCyl),
	nCylBase	:= 12
);

// Desztaplarka - krzywka na falowniku 1
fbSt03.M_ConfigStation(
	pStPersist	:= ADR(GVL_PERSIST.St03),
	pLiftDrive	:= ADR(fbNord[1]),
	nJawId		:= 25,
	pJawPersist	:= ADR(GVL_PERSIST.aCyl[25])
);

// Sztaplarka - falownik krzywki DO USTALENIA.
// Falownik 2 jest na stacji 8, wiec zostaje bez przydzialu.
// Do czasu ustalenia sztaplarka pracuje jako zwykly przelot -
// patrz GVL_PERSIST.aConv[11].Cfg.xStationEnabled ponizej.
fbSt11.M_ConfigStation(
	pStPersist	:= ADR(GVL_PERSIST.St11),
	pLiftDrive	:= 0,
	nJawId		:= 26,
	pJawPersist	:= ADR(GVL_PERSIST.aCyl[26])
);

GVL_PERSIST.aConv[11].Cfg.xStationEnabled := FALSE;


// -------------------------------------------------------------
// LANCUCH TRANSPORTU
// -------------------------------------------------------------
//
// Trasa dobrych:  1 - 2 - 3 - 4 - 5 - 6 - 7 - 8 - 11 - 12 - 13
// Trasa odrzutu:  8 - 9 - 10 - 14 - 15 - 16
// Nastepnik stacji 8 przelacza ACT_Verdict.

fbSt01.M_Link(pPrevNode := 0,            pNextNode := ADR(fbSt02));
fbSt02.M_Link(pPrevNode := ADR(fbSt01),  pNextNode := ADR(fbSt03));
fbSt03.M_Link(pPrevNode := ADR(fbSt02),  pNextNode := ADR(fbSt04));
fbSt04.M_Link(pPrevNode := ADR(fbSt03),  pNextNode := ADR(fbSt05));
fbSt05.M_Link(pPrevNode := ADR(fbSt04),  pNextNode := ADR(fbSt06));
fbSt06.M_Link(pPrevNode := ADR(fbSt05),  pNextNode := ADR(fbSt07));
fbSt07.M_Link(pPrevNode := ADR(fbSt06),  pNextNode := ADR(fbSt08));
fbSt08.M_Link(pPrevNode := ADR(fbSt07),  pNextNode := ADR(fbSt11));

fbSt11.M_Link(pPrevNode := ADR(fbSt08),  pNextNode := ADR(fbSt12));
fbSt12.M_Link(pPrevNode := ADR(fbSt11),  pNextNode := ADR(fbSt13));
fbSt13.M_Link(pPrevNode := ADR(fbSt12),  pNextNode := 0);

fbSt09.M_Link(pPrevNode := ADR(fbSt08),  pNextNode := ADR(fbSt10));
fbSt10.M_Link(pPrevNode := ADR(fbSt09),  pNextNode := ADR(fbSt14));
fbSt14.M_Link(pPrevNode := ADR(fbSt10),  pNextNode := ADR(fbSt15));
fbSt15.M_Link(pPrevNode := ADR(fbSt14),  pNextNode := ADR(fbSt16));
fbSt16.M_Link(pPrevNode := ADR(fbSt15),  pNextNode := 0);
END_ACTION

ACTION ACT_Commands:
// =============================================================
// ACT_Commands
// Komendy operatora
// =============================================================


// -------------------------------------------------------------
// WSTAWIENIE STOSU NA STACJE 1
// -------------------------------------------------------------
//
// Czujnik stacji 1 nie widzi stosu, wiec obecnosc podajemy
// bitem. Stos wjezdza do maszyny jak zwykly ladunek.

rtrgStack(CLK := xCmdStackInserted);

IF rtrgStack.Q THEN

	IF NOT GVL_PERSIST.aConv[1].Mem.xLoadPresent THEN
		nLoadSeq := nLoadSeq + 1;
		fbSt01.M_InjectLoad(xNok := FALSE, nLoadId := nLoadSeq, xOpDone := TRUE);
	END_IF

END_IF


// -------------------------------------------------------------
// KASOWANIE ALARMOW
// -------------------------------------------------------------

rtrgReset(CLK := xCmdReset);

IF rtrgReset.Q THEN
	FOR i := 1 TO 16 DO
		aNode[i]^.M_Reset();
	END_FOR
END_IF


// -------------------------------------------------------------
// RESET MASZYNY DO STANU ZEROWEGO
// -------------------------------------------------------------
//
// Kasuje pamiec obecnosci na wszystkich stacjach oraz liczniki
// desztaplarki i sztaplarki. Uzywac po recznym oproznieniu
// maszyny - maszyna uwierzy, ze jest pusta.

rtrgClear(CLK := xCmdClearMachine);

IF rtrgClear.Q THEN

	FOR i := 1 TO 16 DO
		aNode[i]^.M_ServiceSetEmpty();
	END_FOR

	fbSt03.M_ServiceClearStack();
	fbSt11.M_ServiceClearStack();

	nPalletsDone	:= 0;
	nOkCount		:= 0;
	nNokCount		:= 0;

END_IF
END_ACTION

ACTION ACT_Stations:
// =============================================================
// ACT_Stations
// Wywolanie wszystkich stacji
// =============================================================
//
// Czujniki podajemy w logice WPROST - przelicza je nastawa
// xSensorsInverted w rekordzie stacji.


// Stacja 1 - czujnik nie widzi stosu, wiec pracuje na czasowce
fbSt01(
	eMode			:= eMode,
	xSafetyOK		:= xSafetyOK,
	xTransferEnable	:= xTransferEnable,
	xSens1Raw		:= xSens_St01,
	xSens2Raw		:= FALSE
);

fbSt02(
	eMode			:= eMode,
	xSafetyOK		:= xSafetyOK,
	xTransferEnable	:= xTransferEnable,
	xSens1Raw		:= FALSE,
	xSens2Raw		:= FALSE
);

fbSt03(
	eMode			:= eMode,
	xSafetyOK		:= xSafetyOK,
	xTransferEnable	:= xTransferEnable,
	xSens1Raw		:= xSens_St03,
	xSens2Raw		:= FALSE,
	diLiftPosRaw	:= diEnc_St03,
	xJawClosedSw	:= FALSE,
	xJawOpenSw		:= FALSE
);

// Czujnik wstepny wpisujemy PRZED wywolaniem - inaczej stacja
// zobaczylaby go dopiero w nastepnym cyklu
fbSt04.stIn.xPreSensRaw := xSens_St04_Entry;

fbSt04(
	eMode			:= eMode,
	xSafetyOK		:= xSafetyOK,
	xTransferEnable	:= xTransferEnable,
	xSens1Raw		:= xSens_St04_Stop,
	xSens2Raw		:= FALSE
);

fbSt05(
	eMode			:= eMode,
	xSafetyOK		:= xSafetyOK,
	xTransferEnable	:= xTransferEnable,
	xSens1Raw		:= FALSE,
	xSens2Raw		:= FALSE
);

fbSt06(
	eMode			:= eMode,
	xSafetyOK		:= xSafetyOK,
	xTransferEnable	:= xTransferEnable,
	xSens1Raw		:= FALSE,
	xSens2Raw		:= FALSE
);

fbSt07(
	eMode			:= eMode,
	xSafetyOK		:= xSafetyOK,
	xTransferEnable	:= xTransferEnable,
	xSens1Raw		:= xSens_St07,
	xSens2Raw		:= FALSE
);

fbSt08(
	eMode			:= eMode,
	xSafetyOK		:= xSafetyOK,
	xTransferEnable	:= xTransferEnable,
	xSens1Raw		:= FALSE,
	xSens2Raw		:= FALSE
);

// Transporter lancuchowy - bez wlasnych czujnikow
fbSt09(
	eMode			:= eMode,
	xSafetyOK		:= xSafetyOK,
	xTransferEnable	:= xTransferEnable,
	xSens1Raw		:= FALSE,
	xSens2Raw		:= FALSE
);

fbSt10(
	eMode			:= eMode,
	xSafetyOK		:= xSafetyOK,
	xTransferEnable	:= xTransferEnable,
	xSens1Raw		:= FALSE,
	xSens2Raw		:= FALSE
);

fbSt11(
	eMode			:= eMode,
	xSafetyOK		:= xSafetyOK,
	xTransferEnable	:= xTransferEnable,
	xSens1Raw		:= xSens_St11,
	xSens2Raw		:= FALSE,
	diLiftPosRaw	:= diEnc_St11,
	xJawClosedSw	:= FALSE,
	xJawOpenSw		:= FALSE
);

fbSt12(
	eMode			:= eMode,
	xSafetyOK		:= xSafetyOK,
	xTransferEnable	:= xTransferEnable,
	xSens1Raw		:= FALSE,
	xSens2Raw		:= FALSE
);

fbSt13(
	eMode			:= eMode,
	xSafetyOK		:= xSafetyOK,
	xTransferEnable	:= xTransferEnable,
	xSens1Raw		:= xSens_St13,
	xSens2Raw		:= FALSE,
	xPickupButton	:= FALSE
);

fbSt14(
	eMode			:= eMode,
	xSafetyOK		:= xSafetyOK,
	xTransferEnable	:= xTransferEnable,
	xSens1Raw		:= FALSE,
	xSens2Raw		:= FALSE
);

fbSt15(
	eMode			:= eMode,
	xSafetyOK		:= xSafetyOK,
	xTransferEnable	:= xTransferEnable,
	xSens1Raw		:= FALSE,
	xSens2Raw		:= FALSE
);

fbSt16(
	eMode			:= eMode,
	xSafetyOK		:= xSafetyOK,
	xTransferEnable	:= xTransferEnable,
	xSens1Raw		:= xSens_St16,
	xSens2Raw		:= FALSE,
	xPickupButton	:= FALSE
);


// -------------------------------------------------------------
// CEWKI SZCZEK
// -------------------------------------------------------------

xOut_St03_JawClose	:= fbSt03.xJawCoilClose;
xOut_St03_JawOpen	:= fbSt03.xJawCoilOpen;
xOut_St11_JawClose	:= fbSt11.xJawCoilClose;
xOut_St11_JawOpen	:= fbSt11.xJawCoilOpen;


// -------------------------------------------------------------
// ZAWORY STACJI 4 I 5
// -------------------------------------------------------------

GVL.OUTPUTS[4]	:= fbSt04.stOut.xLowerExtend;
GVL.OUTPUTS[3]	:= fbSt04.stOut.xLowerRetract;
GVL.OUTPUTS[7]	:= fbSt04.stOut.xUpperWideExtend;
GVL.OUTPUTS[2]	:= fbSt04.stOut.xUpperWideRetract;
GVL.OUTPUTS[5]	:= fbSt04.stOut.xUpperNarrowExtend;
GVL.OUTPUTS[6]	:= fbSt04.stOut.xUpperNarrowRetract;

GVL.FestoValves_1[6,1]	:= fbSt05.stOut.xBlockExtend;
GVL.FestoValves_1[6,2]	:= fbSt05.stOut.xBlockRetract;
GVL.FestoValves_1[7,1]	:= fbSt05.stOut.xJawLiftExtend;
GVL.FestoValves_1[7,2]	:= fbSt05.stOut.xJawLiftRetract;

FOR i := 1 TO 3 DO
	GVL.FestoValves_1[i,1] := fbSt05.stOut.axJawClose[i];
END_FOR

// Numer zaworu nie jest numerem silownika - patrz ST_St05_Out
GVL.FestoValves_2[4,2] := fbSt05.stOut.axPullUp[1];
GVL.FestoValves_2[4,1] := fbSt05.stOut.axPullDown[1];
GVL.FestoValves_2[3,2] := fbSt05.stOut.axPullUp[2];
GVL.FestoValves_2[3,1] := fbSt05.stOut.axPullDown[2];
GVL.FestoValves_2[1,2] := fbSt05.stOut.axPullUp[3];
GVL.FestoValves_2[1,1] := fbSt05.stOut.axPullDown[3];
GVL.FestoValves_2[2,2] := fbSt05.stOut.axPullUp[4];
GVL.FestoValves_2[2,1] := fbSt05.stOut.axPullDown[4];
GVL.FestoValves_2[5,2] := fbSt05.stOut.axPullUp[5];
GVL.FestoValves_2[5,1] := fbSt05.stOut.axPullDown[5];
GVL.FestoValves_2[6,2] := fbSt05.stOut.axPullUp[6];
GVL.FestoValves_2[6,1] := fbSt05.stOut.axPullDown[6];
END_ACTION

ACTION ACT_Verdict:
// =============================================================
// ACT_Verdict
// Werdykt OK / NOK oraz trasowanie na stacji 8
// =============================================================
//
// WERSJA TESTOWA. Docelowo werdykt wystawiaja stacje 4, 5 i 6.
// Tutaj co piata paleta idzie na odrzut, zeby przecwiczyc obie
// trasy bez czekania na prawdziwe testy.

rtrgSt05(CLK := GVL_PERSIST.aConv[5].Mem.xOperationDone);

IF rtrgSt05.Q THEN

	nPalletsDone := nPalletsDone + 1;

	IF (nPalletsDone MOD cNokEvery) = 0 THEN
		GVL_PERSIST.aConv[5].Mem.xLoadNok := TRUE;
		nNokCount := nNokCount + 1;
	ELSE
		nOkCount := nOkCount + 1;
	END_IF

END_IF


// -------------------------------------------------------------
// ROZJAZD NA STACJI 8
// -------------------------------------------------------------
//
// Paleta dobra jedzie prosto na sztaplarke, odrzucona
// na transporter poprzeczny.

IF GVL_PERSIST.aConv[8].Mem.xLoadNok THEN
	fbSt08.M_SetNext(pNextNode := ADR(fbSt09));
ELSE
	fbSt08.M_SetNext(pNextNode := ADR(fbSt11));
END_IF
END_ACTION

ACTION ACT_Drives:
// =============================================================
// ACT_Drives
// Wywolanie falownikow - PO stacjach
// =============================================================

FOR i := 1 TO cNumDrives DO

	fbNord[i](
		lrFmax			:= cFmax,
		xSafetyOK		:= xSafetyOK,
		// TODO: podpiac realny status EtherCAT (WcState)
		xEtherCAT_OK	:= TRUE,
		stIn			:= GVL.NORD_DRIVE_IN[i]
	);

	GVL.NORD_DRIVE_OUT[i] := fbNord[i].stOut;

	aeDrvState[i]		:= fbNord[i].eState;
	axDrvRunning[i]		:= fbNord[i].xRunning;
	axDrvError[i]		:= fbNord[i].xError;
	alrDrvFreqAct[i]	:= fbNord[i].lrFreqActual;

END_FOR
END_ACTION

ACTION ACT_Diag:
// =============================================================
// ACT_Diag
// Lustro stanu wszystkich stacji do podgladu online
// =============================================================

FOR i := 1 TO 16 DO
	aeState[i]		:= aNode[i]^.eState;
	aeWait[i]		:= aNode[i]^.eWait;
	aeAlarm[i]		:= aNode[i]^.eAlarm;
	axOccupied[i]	:= aNode[i]^.xOccupied;
	axNok[i]		:= aNode[i]^.xLoadNok;
END_FOR
END_ACTION

END_PROGRAM

// ---- POUs/POUs/FB/TestFb.TcPOU
FUNCTION_BLOCK TestFb
VAR_INPUT
	    stIn            : ST_NordSK550P_In;
END_VAR
VAR_OUTPUT
	    wStatusWord      : UINT;
		dupa2 : INT;
END_VAR
VAR
	dupa : INT := 100;
	i : INT;
END_VAR

wStatusWord := stIn.wStatusWord;
dupa := dupa2;

END_FUNCTION_BLOCK
